// TIA Portal V19 export
TYPE "ST_FieldBus_Output"
   STRUCT
      OUTPUT_BYTE : "ST_Bit";
   END_STRUCT;
END_TYPE
